TYPE ST_JointVelocity :
STRUCT
	q1_dot : LREAL; // dq1 / dt
    q2_dot : LREAL; // dq2 / dt
    q3_dot : LREAL; // dq3 / dt
END_STRUCT
END_TYPE

(* stored: Version 1.1.0.1, ProductVersion 3.1.4024.15
   DUT ST_JointVelocity: Id {574553c2-fc8b-476a-87f3-80f525a49d21} *)
